Fanuc KAREL source: ka00056.KL

PROGRAM KA00056
%STACKSIZE=65535
%PRIORITY=65535
%NOLOCKGROUP
VAR
SRC : POSITION
DST : JOINTPOS9
BEGIN
-- UNSAFE_SOURCE_IR line 7: DST = convert_position_to_jointpos9(SRC)
END KA00056
